Staubli VAL3: actCmd.dtx

public num nMoveID
public num nActionID
public bool bActFinish
public string sActName
